Staubli VAL3: HMI_setting.dtx

mdesc mNomSpeed
bool bBack
bool bMove
bool bTeach
bool bSetup
string sLsit
string sSelTool
string sLastTool
string sList
string sUsingLib
string sLibList
bool bChangeLib
public bool bIsDoing
bool bToSave
bool bLock
bool bDisable[6]
bool bSetMaxJntForce
bool bSix_Axis
string sArmType
num nMaxJntForec[6]
string sArmDetail
string sPassword = "staubli2025"
string sBtnUnLock
